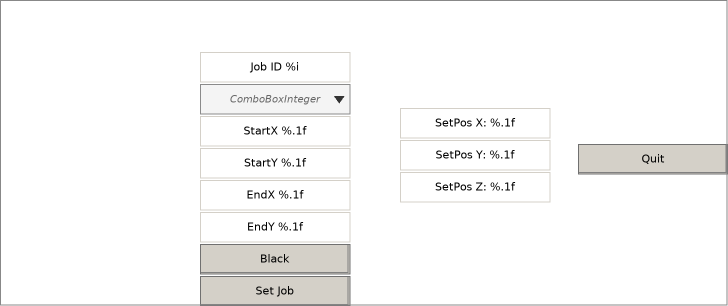
VISUALIZATION VISU  // 728x306
    Textfield (400,108 150x30), "SetPos X: %.1f", text variable: MAIN.fbIgorCtrl.fbPortal.aAxis[X].NcToPlc.SetPos
    Textfield (400,140 150x30), "SetPos Y: %.1f", text variable: MAIN.fbIgorCtrl.fbPortal.aAxis[Y].NcToPlc.SetPos
    Textfield (400,172 150x30), "SetPos Z: %.1f", text variable: MAIN.fbIgorCtrl.fbPortal.aAxis[Z].NcToPlc.SetPos
    Textfield (200,52 150x30), "Job ID %i", text variable: HMI.stJob.nJobID
        OnMouseClick: write HMI.stJob.nJobID via Default
    Textfield (200,180 150x30), "EndX %.1f", text variable: HMI.stJob.fDestPosX
        OnMouseClick: write HMI.stJob.fDestPosX via Default
    Textfield (200,116 150x30), "StartX %.1f", text variable: HMI.stJob.fStartPosX
        OnMouseClick: write HMI.stJob.fStartPosX via Default
    Textfield (200,148 150x30), "StartY %.1f", text variable: HMI.stJob.fStartPosY
        OnMouseClick: write HMI.stJob.fStartPosY via Default
    Textfield (200,212 150x30), "EndY %.1f", text variable: HMI.stJob.fDestPosY
        OnMouseClick: write HMI.stJob.fDestPosY via Default
    Button (200,276 150x30), "Set Job"
        tap HMI.bSetJob
    Button (578,144 150x30), "Quit"
        tap HMI.bQuit
    ComboBoxInteger (200,84 150x30), variable: HMI.stJob.eJobType
    Button (200,244 150x30), "Black"
        toggle HMI.stJob.bBlack
END_VISUALIZATION

(* stored: Version 1.1.0.1, ProductVersion 3.1.4024.9
   Visu VISU: Id {9cb3c082-dce7-4ea0-924b-7993a5243e75} *)
